(* IEC 61131-3 sources: codesys-to-astra/tests/POUs/FB_C2aTime_Test, 6 files *)

(* ---- FB_C2aTime_Test.decl.st ---- *)
// Назначение: тесты календаря F_C2aUnixToDate и форматов FB_C2aRtc (ожидания — по календарю, не по коду).
// Автор:      kr0nsch
// Версия:     0.1.0
// Документ:   docs/TEST_REPORT.md
FUNCTION_BLOCK FB_C2aTime_Test EXTENDS coUnit.FB_TestSuite
VAR CONSTANT
    R_DELTA : REAL := 0.0001;   // допуск сравнения REAL
END_VAR

(* ---- Epoch.method.decl.st ---- *)
// 0 -> 1970-01-01 00:00:00, четверг (4)
METHOD PRIVATE Epoch
VAR
    stD : ST_C2aDateTime;  // результат
END_VAR

(* ---- LeapDay.method.decl.st ---- *)
// 951782400 -> 2000-02-29 00:00:00, вторник (2)
METHOD PRIVATE LeapDay
VAR
    stD : ST_C2aDateTime;  // результат
END_VAR

(* ---- Pad2.method.decl.st ---- *)
// F_C2aPad2: 7 -> '07', 42 -> '42'
METHOD PRIVATE Pad2
VAR
    s7 : STRING(2);  // 7
    s42 : STRING(2);  // 42
END_VAR

(* ---- RtcReadsClock.method.decl.st ---- *)
// FB_C2aRtc читает часы рантайма: год не меньше 2024, xOk
METHOD PRIVATE RtcReadsClock
VAR
    fbRtc : FB_C2aRtc;  // время рантайма
END_VAR

(* ---- TimeOfDay.method.decl.st ---- *)
// 1792494245 -> 2026-10-20 11:04:05, вторник
METHOD PRIVATE TimeOfDay
VAR
    stD : ST_C2aDateTime;  // результат
END_VAR
